(* IEC 61131-3 sources: PortalRobot/Portal_robot/Device/application/FB (part 4) *)

(* ---- FB_MAGAZINE.st ---- *)
FUNCTION_BLOCK FB_MAGAZINE
VAR_INPUT
	xIoManual : BOOL; // Передача выходов оператору отменяет пошаговую операцию
	uiMagazineId : UINT; // Идентификатор экземпляра 1..2
	xPointsConfigured : BOOL; // Настроена база этого магазина с Safe Z и Change Z
	xMechanismReady : BOOL := TRUE;
	xInventoryChanged : BOOL; // Сменился рабочий банк или оператор изменил его содержимое
	xTestInitialize : BOOL;
	xTestEnabled : BOOL;
	stRobotStatus     : ST_ROBOT_STATUS; // Текущие статусы робота
	astMachineStatus  : ARRAY [1..3] OF ST_MACHINE_PUBLIC; // Статусы станков для определения оставшейся работы
	auiMachineType    : ARRAY [1..3] OF UINT; // Тип детали, закреплённый за каждым станком
	stMagazineCommand : ST_MAGAZINE_COMMAND; // Команда магазина от автоматической логики
	stHmiCommand      : ST_ROBOT_COMMAND; // Ручная команда магазина с HMI
	xManual           : BOOL; // Разрешение ручного управления
	xReset            : BOOL; // Сброс ошибок магазина
	xResetCancel      : BOOL; // Отмена согласованного сброса по Stop/Disable
	RobotResetRecovery : ST_ROBOT_RESET_RECOVERY; // Внутреннее подтверждение принятого Reset робота
	xGlobalError      : BOOL; // Глобальная ошибка ячейки
	xHmiEnable        : BOOL; // Импульс включения магазина с HMI
	xHmiDisable       : BOOL; // Импульс отключения магазина с HMI
	xHmiFillBlanks    : BOOL; // Заполнить все активные слоты матрицы заготовками
	xHmiClear         : BOOL; // Полностью очистить содержимое магазина
	xHmiCycleSlot     : BOOL; // Переключить содержимое выбранного слота
	xHmiApplySlot     : BOOL; // Явно записать состояние и тип выбранного слота
	xHmiApplyPitchX   : BOOL; // Применить новый общий шаг слотов по X
	xHmiApplyPitchY   : BOOL; // Применить новый общий шаг слотов по Y
	uiHmiEditSlot     : UINT; // Номер слота для ручного редактирования
	uiHmiEditDetailType : UINT; // 0=NONE, 1=BLANK, 2=DETAIL
	uiHmiEditProductType : UINT; // Тип изделия 1..3
	lrHmiEditPitchX   : LREAL;
	lrHmiEditPitchY   : LREAL;
	xRobotOwnsMagazine : BOOL; // Автомат удерживает этот магазин в текущем цикле
	xRobotCanWorkWithMagazine : BOOL; // Интерфейс и точки готовы для роботной операции, не для включения магазина
	xSharedGeometryEditAllowed : BOOL; // Оба магазина выключены; общий шаг можно менять
	uiRows            : UINT; // Число строк матрицы магазина
	uiColumns         : UINT; // Число столбцов матрицы магазина
	uiTypeCount       : UINT; // Количество настроенных типов заготовок, 1..3
	auiSlotType       : ARRAY [1..GVL_CELL_SETTINGS.NumberDetail] OF UINT; // Тип секции каждого слота
	FaultRequest  : ST_MAGAZINE_FAULT_REQUEST; // Единый контракт диагностической инъекции
END_VAR
VAR_OUTPUT
    xInventoryUpdated : BOOL; // Только записи содержимого этим FB в текущем скане
	Command : ST_ROBOT_COMMAND; // Текущая пошаговая команда роботу
	Status  : ST_MAGAZINE_STATUS; // Рабочие статусы магазина
	Diag    : ST_MAGAZINE_DIAG; // Состояние автомата магазина
	Error   : ST_MAGAZINE_ERRORS; // Активные и последние ошибки
	FaultStatus : ST_FAULT_INJECTION_STATUS; // Состояние инжектора для HMI
END_VAR
VAR_IN_OUT
	stInventory : ST_MAGAZINE_INVENTORY; // Единственная кассета текущего магазина
	lrPitchX : LREAL; // Общий фактический шаг слотов по X
	lrPitchY : LREAL; // Общий фактический шаг слотов по Y
END_VAR
VAR
    xInventorySummaryInitialized : BOOL;
    xInventorySummaryDirty : BOOL;
    iInventorySummarySlotCount : SINT;
    uiInventorySummaryTypeCount : UINT;
    iInventoryFirstBlank : SINT;
    iInventoryFirstFree : SINT;
	eGrantedOperation : E_MAGAZINE_OPERATION; // Доступная операция магазина
	eActualOperation  : E_MAGAZINE_OPERATION; // Выполняемая операция магазина

	rtExecute          : R_TRIG; // Фронт команды запуска
	rtEnable           : R_TRIG; // Фронт команды включения
	rtDisable          : R_TRIG; // Фронт команды отключения
	rtFillBlanks       : R_TRIG; // Фронт заполнения магазина заготовками
	rtClear            : R_TRIG; // Фронт очистки магазина
	rtCycleSlot        : R_TRIG; // Фронт изменения выбранного слота
	rtApplySlot        : R_TRIG; // Фронт явной записи выбранного слота
	rtApplyPitchX      : R_TRIG;
	rtApplyPitchY      : R_TRIG;
	rtReset            : R_TRIG; // Фронт команды сброса магазина

	xExecuteRequest    : BOOL; // Активный запрос выполнения операции
	xResetRequest      : BOOL; // Активный запрос сброса
	xStopRequest       : BOOL; // Активный запрос остановки
	xManualCommand     : BOOL; // Команда получена из ручного интерфейса
	xDisableRequest    : BOOL; // Сохранённый запрос отключения после текущей операции
	xRobotInMagazineContext : BOOL; // Робот находится в рабочей зоне магазина
	xFaultContextCaptured : BOOL; // Контекст робота зафиксирован при входе в ERROR
	xRobotInMagazineAtFault : BOOL; // Робот был в рабочей зоне этого магазина при ошибке
	xRobotStopRequired : BOOL; // Итоговая реакция ROBOT_STOP, сформированная магазином
	xRobotResetDependencyReady : BOOL; // Каскадная ошибка робота может быть сброшена тем же импульсом
	xRobotResetDependencyRequired : BOOL; // Только ошибка с участием робота зависит от его восстановления
	xRobotResetCoordinated : BOOL; // Магазин присоединился к одному явно запрошенному сбросу
	udiRobotResetAttempt : UDINT; // Ожидаемый номер принятой попытки FB_ROBOT
	xRobotResetAttemptReady : BOOL; // Первичная зависимость восстановлена в той же попытке

	iActiveSlotCount   : SINT; // Число активных слотов выбранной матрицы
	iInventoryIndex    : SINT; // Индекс изменения содержимого магазина
	iTakeSlot          : SINT; // Слот выбранной заготовки
	iPutSlot           : SINT; // Выбранный свободный слот
	iActiveSlot        : SINT; // Единственный слот текущего элементарного движения
	xInventoryCommitted: BOOL; // Все изменения слотов текущей операции подтверждены
	xTakeSlotCommitted  : BOOL; // Изъятие заготовки отражено в матрице после закрытия захвата
	xPutSlotCommitted   : BOOL; // Укладка груза отражена в матрице после открытия захвата
	xRobotCommandStarted : BOOL; // Текущий элементарный шаг действительно принят FB_ROBOT
	xOperationSequenceComplete : BOOL; // Все шаги операции подтверждены до изменения матрицы
	xTakeSlotValid     : BOOL; // Проверка диапазона до обращения к массиву слотов
	xPutSlotValid      : BOOL;
	xTakeSlotHasBlank  : BOOL;
	xPutSlotEmpty      : BOOL;
	xChangeTakeFirst   : BOOL; // CHANGE в одном слоте: сначала TAKE, затем PUT
	xPutProductTypeValid : BOOL;
	uiStep             : UINT; // Шаг последовательности робота
	uiIndex            : UINT; // Индекс слота для расчёта координат

	stActiveRobotCommand : ST_ROBOT_COMMAND; // Команда роботу текущего шага
	xFinishedCondition   : BOOL; // Текущее содержимое не позволяет продолжить цикл
	xFinishedLatched     : BOOL; // Завершение этой палеты не отменяется работой другого магазина
	xMachineHasRelevantPart : BOOL; // В доступном станке есть заготовка, обработка или готовая деталь
	xMachineHasDestination : BOOL; // Для оставшейся работы есть свободный слот соответствующего типа
	xAllSlotsDetails    : BOOL; // Все активные слоты заполнены готовыми деталями
	xNoBlankNoMachinePart : BOOL; // Нет заготовок и нет доступной работы в станках
	xNoBlankNoDestination : BOOL; // Нет заготовок и нет места для возврата груза
	uiMachineIndex      : UINT; // Индекс станка при расчёте завершения магазина
	uiMachineTypeIndex  : UINT; // Тип детали проверяемого станка
	uiPutProductType    : UINT; // Тип груза, защёлкнутый до физического PUT
	fbFaultInjector      : FB_MAGAZINE_FAULT_INJECTOR; // Безопасный сценарий ошибки до движения
	xFaultAllowed        : BOOL; // Владелец разрешает синтетическую проверку
	xStartupInitialized  : BOOL;
	udiProducedPartsTotal : UDINT; // Монотонный счётчик подтверждённых укладок готовых деталей
END_VAR
VAR CONSTANT
	ERR_WRONG_OPERATION : DWORD := DWORD#16#0000_0001; // Недопустимая операция магазина
	ERR_NO_BLANK        : DWORD := DWORD#16#0000_0002; // В магазине нет заготовки
	ERR_NO_FREE_SLOT    : DWORD := DWORD#16#0000_0004; // В магазине нет свободного слота
	ERR_INVALID_SLOT    : DWORD := DWORD#16#0000_0008; // Недопустимый номер слота
	ERR_SLOT_CONTENT    : DWORD := DWORD#16#0000_0010; // Содержимое слота не соответствует операции
	ERR_ROBOT           : DWORD := DWORD#16#0000_0020; // Ошибка робота при операции магазина
	ERR_GLOBAL_STOP     : DWORD := DWORD#16#0000_0040; // Остановка по глобальной ошибке
	ERR_GEOMETRY        : DWORD := DWORD#16#0000_0080; // Ошибка параметров матрицы магазина
	MASK_EQUIPMENT_ERROR : DWORD := ERR_WRONG_OPERATION OR ERR_NO_BLANK
		OR ERR_NO_FREE_SLOT OR ERR_INVALID_SLOT OR ERR_SLOT_CONTENT OR ERR_GEOMETRY;
	WRN_RESET_EXECUTE_ACTIVE : UINT := 1; // Операция магазина ещё активна
	WRN_RESET_GLOBAL_ERROR   : UINT := 2; // Глобальная ошибка ещё активна
	WRN_RESET_ROBOT_ERROR    : UINT := 3; // Ошибка робота ещё активна
	WRN_ENABLE_GLOBAL_ERROR  : UINT := 4; // Включение запрещено глобальной ошибкой
	WRN_ENABLE_CONTENT       : UINT := 5; // Архив: содержимое больше не блокирует включение
	WRN_DISABLE_PENDING      : UINT := 6; // Отключение магазина уже запрошено
	WRN_FILL_ENABLED         : UINT := 7; // Заполнение запрещено для включённого магазина
	WRN_FILL_GEOMETRY        : UINT := 8; // Активная матрица магазина задана неверно
	WRN_CLEAR_ENABLED        : UINT := 9; // Очистка запрещена для включённого магазина
	WRN_SIM_ERROR_NOT_ALLOWED: UINT := 10; // Тестовая ошибка запрещена текущим состоянием
	WRN_EDIT_REJECTED : UINT := 14; // Редактирование включённого/занятого магазина запрещено
	WRN_GEOMETRY_EDIT_REJECTED : UINT := 16; // PLC отклонил изменение общего шага X/Y
	WRN_ENABLE_GEOMETRY      : UINT := 15; // Геометрия магазина не позволяет включение
	WRN_ENABLE_OWN_ERROR     : UINT := 17; // Включение запрещено собственной ошибкой магазина
	WRN_ENABLE_POINTS        : UINT := 18; // Не настроена база этого магазина или её Z-смещения
END_VAR

// --- BEGIN IMPLEMENTATION ---

xInventoryUpdated := FALSE;

// Инвентарь загружает владелец банков RunTwoPallet; здесь сбрасывается только автомат.
IF NOT xStartupInitialized THEN
	xFinishedLatched := FALSE;
	xFaultContextCaptured := FALSE;
	xRobotInMagazineAtFault := FALSE;
	xRobotStopRequired := FALSE;
	xStartupInitialized := TRUE;
END_IF;

IF xTestInitialize THEN
	xFinishedLatched := FALSE;
	IF xTestEnabled AND xPointsConfigured THEN
		Diag.eState := E_MAGAZINE_STATE.IDLE;
	ELSE
		Diag.eState := E_MAGAZINE_STATE.DISABLED;
	END_IF;
	Error.dwErrorActive := DWORD#0;
	Error.dwAlarmActive := DWORD#0;
	eGrantedOperation := E_MAGAZINE_OPERATION.NONE;
	eActualOperation := E_MAGAZINE_OPERATION.NONE;
	xExecuteRequest := FALSE;
	xResetRequest := FALSE;
	xStopRequest := FALSE;
	xManualCommand := FALSE;
	xDisableRequest := FALSE;
	iTakeSlot := SINT#0;
	iPutSlot := SINT#0;
	xChangeTakeFirst := FALSE;
	iActiveSlot := SINT#0;
	xInventoryCommitted := FALSE;
	xTakeSlotCommitted := FALSE;
	xPutSlotCommitted := FALSE;
	xRobotCommandStarted := FALSE;
	xOperationSequenceComplete := FALSE;
	xFaultContextCaptured := FALSE;
	xRobotInMagazineAtFault := FALSE;
	xRobotStopRequired := FALSE;
	uiStep := UINT#0;
	stActiveRobotCommand.xExecute := FALSE;
	stActiveRobotCommand.xStop := FALSE;
	stActiveRobotCommand.xReset := FALSE;
	stActiveRobotCommand.eAction := E_ROBOT_ACTION.NONE;
	stActiveRobotCommand.eSetPoint := E_POINT_NAME.NONE;
	stActiveRobotCommand.iActiveSlot := SINT#0;
	stActiveRobotCommand.uiMagazineId := uiMagazineId;
END_IF;

IF xInventoryChanged THEN
	xFinishedLatched := FALSE;
END_IF;

rtFillBlanks(CLK := xHmiFillBlanks);
rtClear(CLK := xHmiClear);
rtCycleSlot(CLK := xHmiCycleSlot);
rtApplySlot(CLK := xHmiApplySlot);
rtApplyPitchX(CLK := xHmiApplyPitchX);
rtApplyPitchY(CLK := xHmiApplyPitchY);

IF (uiRows > UINT#0)
AND (uiColumns > UINT#0)
AND ((uiRows * uiColumns) <= SINT_TO_UINT(GVL_CELL_SETTINGS.MagazineSlots)) THEN
	iActiveSlotCount := UINT_TO_SINT(uiRows * uiColumns);
ELSE
	iActiveSlotCount := SINT#0;
END_IF;

// Ручная роботная команда принадлежит только выбранному магазину.
xManualCommand := xManual
	AND (
		(stHmiCommand.eSetPoint = E_POINT_NAME.MAGAZINE_TAKE_DETAIL)
		OR (stHmiCommand.eSetPoint = E_POINT_NAME.MAGAZINE_PUT_DETAIL)
		OR (stHmiCommand.eSetPoint = E_POINT_NAME.MAGAZINE_CHANGE_DETAIL)
		OR (stHmiCommand.eSetPoint = E_POINT_NAME.MAGAZINE_RETURN_BLANK)
	)
	AND ((stHmiCommand.uiMagazineId = uiMagazineId)
		OR ((stHmiCommand.uiMagazineId = UINT#0) AND (uiMagazineId = UINT#1)));

IF xManual THEN
	IF xManualCommand THEN
		xExecuteRequest := stHmiCommand.xExecute;
		xStopRequest := stHmiCommand.xStop;
	ELSE
		xExecuteRequest := FALSE;
		xStopRequest := FALSE;
	END_IF;
ELSE
	xExecuteRequest := stMagazineCommand.xExecute;
	xStopRequest := stMagazineCommand.xStop;
END_IF;

// Контекст запрещает редактирование и завершает отложенное отключение только
// после фактического выхода робота из конкретного магазина.
xRobotInMagazineContext := (stRobotStatus.uiMagazineContext = uiMagazineId)
	OR ((stRobotStatus.uiMagazineContext = UINT#0)
		AND (xRobotOwnsMagazine OR xManualCommand)
		AND ((stRobotStatus.eCurrentPoint = E_POINT_NAME.MAGAZINE_IN_SLOT)
			OR (stRobotStatus.eCurrentPoint = E_POINT_NAME.MAGAZINE_CHANGE)));
xRobotInMagazineContext := xRobotInMagazineContext
	OR ((xRobotOwnsMagazine OR xManualCommand)
		AND (Diag.eState = E_MAGAZINE_STATE.ROBOT_COMMAND)
		AND (stActiveRobotCommand.eAction = E_ROBOT_ACTION.MOVE_TO_POINT)
		AND ((stActiveRobotCommand.eSetPoint = E_POINT_NAME.MAGAZINE_IN_SLOT)
			OR (stActiveRobotCommand.eSetPoint = E_POINT_NAME.MAGAZINE_CHANGE)));

// Единственную кассету можно менять только у технологически выключенного
// магазина, когда робот не находится внутри и не владеет текущей операцией.
Status.xEditAllowed := ((Diag.eState = E_MAGAZINE_STATE.DISABLED)
		OR (Diag.eState = E_MAGAZINE_STATE.ERROR))
	AND NOT xRobotOwnsMagazine
	AND NOT xRobotInMagazineContext
	AND NOT xGlobalError;
Status.xPitchEditAllowed := Status.xEditAllowed AND xSharedGeometryEditAllowed;

// Шаг матрицы общий для двух магазинов, поэтому менять его разрешено только
// когда оба магазина выключены. Смещения Z принадлежат базовым точкам магазина.
IF rtApplyPitchX.Q
AND Status.xEditAllowed
AND xSharedGeometryEditAllowed
AND (lrHmiEditPitchX >= LREAL#1.0)
AND (lrHmiEditPitchX <= LREAL#5000.0) THEN
	lrPitchX := lrHmiEditPitchX;
END_IF;
IF rtApplyPitchY.Q
AND Status.xEditAllowed
AND xSharedGeometryEditAllowed
AND (lrHmiEditPitchY >= LREAL#1.0)
AND (lrHmiEditPitchY <= LREAL#5000.0) THEN
	lrPitchY := lrHmiEditPitchY;
END_IF;
IF rtClear.Q AND Status.xEditAllowed THEN
	xFinishedLatched := FALSE;
	FOR iInventoryIndex := 1 TO GVL_CELL_SETTINGS.MagazineSlots DO
		xInventoryUpdated := TRUE;
		xInventorySummaryDirty := TRUE;
		stInventory.aSlots[iInventoryIndex].xInPosition := FALSE;
		stInventory.aSlots[iInventoryIndex].eDetailType := E_DETAIL_TYPE.NONE;
		stInventory.aSlots[iInventoryIndex].uiProductType := UINT#0;
	END_FOR;
ELSIF rtFillBlanks.Q
AND (iActiveSlotCount > SINT#0)
AND Status.xEditAllowed THEN
	xFinishedLatched := FALSE;
	FOR iInventoryIndex := 1 TO GVL_CELL_SETTINGS.MagazineSlots DO
		xInventoryUpdated := TRUE;
		xInventorySummaryDirty := TRUE;
		stInventory.aSlots[iInventoryIndex].xInPosition := iInventoryIndex <= iActiveSlotCount;
		IF iInventoryIndex <= iActiveSlotCount THEN
			stInventory.aSlots[iInventoryIndex].eDetailType := E_DETAIL_TYPE.BLANK;
			stInventory.aSlots[iInventoryIndex].uiProductType := auiSlotType[iInventoryIndex];
		ELSE
			stInventory.aSlots[iInventoryIndex].eDetailType := E_DETAIL_TYPE.NONE;
			stInventory.aSlots[iInventoryIndex].uiProductType := UINT#0;
		END_IF;
	END_FOR;
ELSIF rtApplySlot.Q
AND Status.xEditAllowed
AND (uiHmiEditSlot >= UINT#1)
AND (uiHmiEditSlot <= SINT_TO_UINT(iActiveSlotCount))
AND (uiHmiEditDetailType <= UINT#2)
AND ((uiHmiEditDetailType = UINT#0)
	OR ((uiHmiEditProductType >= UINT#1) AND (uiHmiEditProductType <= uiTypeCount))) THEN
	xFinishedLatched := FALSE;
	iInventoryIndex := UINT_TO_SINT(uiHmiEditSlot);
	CASE uiHmiEditDetailType OF
		UINT#0:
			xInventoryUpdated := TRUE;
			xInventorySummaryDirty := TRUE;
			stInventory.aSlots[iInventoryIndex].xInPosition := FALSE;
			stInventory.aSlots[iInventoryIndex].eDetailType := E_DETAIL_TYPE.NONE;
			stInventory.aSlots[iInventoryIndex].uiProductType := UINT#0;
		UINT#1:
			xInventoryUpdated := TRUE;
			xInventorySummaryDirty := TRUE;
			stInventory.aSlots[iInventoryIndex].xInPosition := TRUE;
			stInventory.aSlots[iInventoryIndex].eDetailType := E_DETAIL_TYPE.BLANK;
			stInventory.aSlots[iInventoryIndex].uiProductType := uiHmiEditProductType;
		UINT#2:
			xInventoryUpdated := TRUE;
			xInventorySummaryDirty := TRUE;
			stInventory.aSlots[iInventoryIndex].xInPosition := TRUE;
			stInventory.aSlots[iInventoryIndex].eDetailType := E_DETAIL_TYPE.DETAIL;
			stInventory.aSlots[iInventoryIndex].uiProductType := uiHmiEditProductType;
	END_CASE;
ELSIF rtCycleSlot.Q
AND Status.xEditAllowed
AND (uiHmiEditSlot >= UINT#1)
AND (uiHmiEditSlot <= SINT_TO_UINT(iActiveSlotCount)) THEN
	xFinishedLatched := FALSE;
	iInventoryIndex := UINT_TO_SINT(uiHmiEditSlot);
	IF NOT stInventory.aSlots[iInventoryIndex].xInPosition
	OR (stInventory.aSlots[iInventoryIndex].eDetailType = E_DETAIL_TYPE.NONE) THEN
		xInventoryUpdated := TRUE;
		xInventorySummaryDirty := TRUE;
		stInventory.aSlots[iInventoryIndex].xInPosition := TRUE;
		stInventory.aSlots[iInventoryIndex].eDetailType := E_DETAIL_TYPE.BLANK;
		stInventory.aSlots[iInventoryIndex].uiProductType := auiSlotType[iInventoryIndex];
	ELSE
		xInventoryUpdated := TRUE;
		xInventorySummaryDirty := TRUE;
		stInventory.aSlots[iInventoryIndex].xInPosition := FALSE;
		stInventory.aSlots[iInventoryIndex].eDetailType := E_DETAIL_TYPE.NONE;
		stInventory.aSlots[iInventoryIndex].uiProductType := UINT#0;
	END_IF;
END_IF;

// При смене банка проверка завершения использует его текущую карту типов,
// а не свободные слоты прежней палеты с прошлого скана.
IF NOT xInventorySummaryInitialized OR xInventoryChanged OR xTestInitialize
OR (iInventorySummarySlotCount <> iActiveSlotCount)
OR (uiInventorySummaryTypeCount <> uiTypeCount) THEN
    xInventorySummaryDirty := TRUE;
END_IF;
IF xInventorySummaryDirty THEN
    UpdateTypeStatus(stMagazineInventory := stInventory);
END_IF;
Status.iCurrentBlank := iInventoryFirstBlank;
Status.iCurrentFreeSlot := iInventoryFirstFree;

Status.xOutBlank := Status.iCurrentBlank = SINT#0;
Status.xOutFreeSlot := Status.iCurrentFreeSlot = SINT#0;
Status.xCanTake := NOT Status.xOutBlank;
Status.xCanPut := NOT Status.xOutFreeSlot;
Status.xCanChange := Status.xCanTake; // Изъятие заготовки само освобождает место
Status.xCanEnable := FALSE;

// Для PUT/возврата заготовки нужен пустой слот. Готовую деталь можно обменять
// на заготовку в одном занятом слоте, если первый захват свободен и открыт.
IF stRobotStatus.xBlankAvailable OR stRobotStatus.xDetailAvailable THEN
	Status.xCanEnable := Status.xCanPut;
ELSIF NOT stRobotStatus.xBlankAvailable AND NOT stRobotStatus.xDetailAvailable THEN
	Status.xCanEnable := Status.xCanTake;
END_IF;

IF stRobotStatus.xDetailAvailable AND NOT stRobotStatus.xBlankAvailable
AND stRobotStatus.xGripper1Open AND Status.xCanChange THEN
	Status.xCanEnable := TRUE;
END_IF;

// Отсутствие заготовок не завершает магазин, пока из станков ещё можно вернуть
// готовую деталь в свободный слот соответствующего типа.
xMachineHasRelevantPart := FALSE;
xMachineHasDestination := FALSE;
FOR uiMachineIndex := UINT#1 TO UINT#3 DO
	IF astMachineStatus[uiMachineIndex].xEnabled
	AND NOT astMachineStatus[uiMachineIndex].xError
	AND (astMachineStatus[uiMachineIndex].xProcessing
		OR ((astMachineStatus[uiMachineIndex].ePartState = E_PART_STATE.LOADED)
			AND ((astMachineStatus[uiMachineIndex].ePartType = E_PART_TYPE.PART)
				OR (astMachineStatus[uiMachineIndex].ePartType = E_PART_TYPE.DETAIL)))) THEN
		xMachineHasRelevantPart := TRUE;
		uiMachineTypeIndex := auiMachineType[uiMachineIndex];
		IF (uiMachineTypeIndex >= UINT#1)
		AND (uiMachineTypeIndex <= UINT#3)
		AND (Status.stTypeStatus.aiFreeSlot[uiMachineTypeIndex] > SINT#0) THEN
			xMachineHasDestination := TRUE;
		END_IF;
	END_IF;
END_FOR;

IF NOT stRobotStatus.xBlankAvailable
AND NOT stRobotStatus.xDetailAvailable
AND xMachineHasDestination THEN
	Status.xCanEnable := TRUE;
END_IF;

Status.xEnableCheckRobotReady := xRobotCanWorkWithMagazine AND xMechanismReady;
Status.xEnableCheckRobotReleased := NOT xRobotInMagazineContext;
Status.xEnableCheckNoError := NOT xGlobalError
	AND (Diag.eState <> E_MAGAZINE_STATE.ERROR)
	AND (Error.dwErrorActive = DWORD#0);
Status.xEnableCheckContent := Status.xCanEnable;
Status.xEnableCheckGeometry := (iActiveSlotCount > SINT#0)
	AND (lrPitchX >= LREAL#1.0)
	AND (lrPitchX <= LREAL#5000.0)
	AND (lrPitchY >= LREAL#1.0)
	AND (lrPitchY <= LREAL#5000.0);
// Включение требует собственную базовую точку магазина. Готовность интерфейса,
// положение робота и содержимое палеты проверяются при роботной операции.
Status.xEnableSequenceAllowed := (Diag.eState = E_MAGAZINE_STATE.DISABLED)
	AND Status.xEnableCheckNoError
	AND Status.xEnableCheckGeometry
	AND xPointsConfigured;

// Finished остаётся прежним по смыслу, но теперь оценивает единственную кассету.
xAllSlotsDetails := iActiveSlotCount > SINT#0;
IF xAllSlotsDetails THEN
	FOR uiIndex := UINT#1 TO SINT_TO_UINT(iActiveSlotCount) DO
		IF NOT stInventory.aSlots[UINT_TO_SINT(uiIndex)].xInPosition
		OR (stInventory.aSlots[UINT_TO_SINT(uiIndex)].eDetailType <> E_DETAIL_TYPE.DETAIL) THEN
			xAllSlotsDetails := FALSE;
		END_IF;
	END_FOR;
END_IF;
xNoBlankNoMachinePart := Status.xOutBlank AND NOT xMachineHasRelevantPart;
xNoBlankNoDestination := Status.xOutBlank AND NOT xMachineHasDestination;
xFinishedCondition :=
	(NOT stRobotStatus.xBlankAvailable AND NOT stRobotStatus.xDetailAvailable)
	AND (xAllSlotsDetails OR xNoBlankNoMachinePart OR xNoBlankNoDestination);

eGrantedOperation := E_MAGAZINE_OPERATION.NONE;
IF stRobotStatus.xBlankAvailable
AND stRobotStatus.xDetailAvailable
AND Status.xCanPut THEN
	// Сначала освобождается захват готовой детали; заготовка остаётся у робота.
	eGrantedOperation := E_MAGAZINE_OPERATION.PUT;
ELSIF NOT Status.xOutBlank
AND NOT stRobotStatus.xBlankAvailable
AND NOT stRobotStatus.xDetailAvailable THEN
	eGrantedOperation := E_MAGAZINE_OPERATION.TAKE;
ELSIF NOT Status.xOutBlank
AND stRobotStatus.xGripper1Open
AND NOT stRobotStatus.xBlankAvailable
AND stRobotStatus.xDetailAvailable THEN
	eGrantedOperation := E_MAGAZINE_OPERATION.CHANGE;
ELSIF NOT Status.xOutFreeSlot
AND stRobotStatus.xDetailAvailable THEN
	eGrantedOperation := E_MAGAZINE_OPERATION.PUT;
END_IF;

xResetRequest := xReset;
rtReset(CLK := xResetRequest);

// RunMagazine предшествует RunRobot. В скане нажатия ожидаем следующий номер;
// на следующем скане уже требуется подтверждённая, всё ещё активная попытка.
IF xRobotResetCoordinated
AND (NOT RobotResetRecovery.xActive
	OR (RobotResetRecovery.udiAttempt <> udiRobotResetAttempt)
	OR xGlobalError OR xIoManual OR xStopRequest OR xExecuteRequest OR xResetCancel) THEN
	xRobotResetCoordinated := FALSE;
	IF (Diag.eState = E_MAGAZINE_STATE.ERROR) AND stRobotStatus.xError THEN
		Diag.stWarning.uiCode := WRN_RESET_ROBOT_ERROR;
		Diag.stWarning.udiSequence := Diag.stWarning.udiSequence + UDINT#1;
		IF Diag.stWarning.udiSequence = UDINT#0 THEN Diag.stWarning.udiSequence := UDINT#1; END_IF;
	END_IF;
END_IF;
xRobotResetAttemptReady := xRobotResetCoordinated
	AND RobotResetRecovery.xActive
	AND (RobotResetRecovery.udiAttempt = udiRobotResetAttempt)
	AND RobotResetRecovery.xDependenciesReady;

xRobotResetDependencyRequired := ((Error.dwErrorActive AND ERR_ROBOT) <> DWORD#0)
	OR xRobotInMagazineAtFault;
xRobotResetDependencyReady := NOT xRobotResetDependencyRequired
	OR NOT stRobotStatus.xError
	OR stRobotStatus.xResetAllowed
	OR xRobotResetAttemptReady;

IF rtReset.Q
AND (Diag.eState = E_MAGAZINE_STATE.ERROR) THEN
	IF xExecuteRequest THEN
		Diag.stWarning.uiCode := WRN_RESET_EXECUTE_ACTIVE;
	ELSIF xGlobalError THEN
		Diag.stWarning.uiCode := WRN_RESET_GLOBAL_ERROR;
	ELSIF stRobotStatus.xError
	AND NOT stRobotStatus.xResetAllowed THEN
		Diag.stWarning.uiCode := WRN_RESET_ROBOT_ERROR;
	ELSE
		Diag.stWarning.uiCode := UINT#0;
	END_IF;

	IF Diag.stWarning.uiCode <> UINT#0 THEN
		Diag.stWarning.udiSequence := Diag.stWarning.udiSequence + UDINT#1;
		IF Diag.stWarning.udiSequence = UDINT#0 THEN
			Diag.stWarning.udiSequence := UDINT#1;
		END_IF;
	END_IF;
END_IF;

rtEnable(CLK := xHmiEnable OR (NOT xManual AND stMagazineCommand.xEnable));
rtDisable(CLK := xHmiDisable OR (NOT xManual AND stMagazineCommand.xDisable));

IF rtEnable.Q
AND (Diag.eState = E_MAGAZINE_STATE.DISABLED)
AND NOT Status.xEnableSequenceAllowed THEN
	IF NOT xPointsConfigured THEN
		Diag.stWarning.uiCode := WRN_ENABLE_POINTS;
	ELSIF xGlobalError THEN
		Diag.stWarning.uiCode := WRN_ENABLE_GLOBAL_ERROR;
	ELSIF NOT Status.xEnableCheckGeometry THEN
		Diag.stWarning.uiCode := WRN_ENABLE_GEOMETRY;
	ELSE
		Diag.stWarning.uiCode := WRN_ENABLE_OWN_ERROR;
	END_IF;
	Diag.stWarning.udiSequence := Diag.stWarning.udiSequence + UDINT#1;
	IF Diag.stWarning.udiSequence = UDINT#0 THEN
		Diag.stWarning.udiSequence := UDINT#1;
	END_IF;
ELSIF rtDisable.Q
AND xHmiDisable
AND xDisableRequest THEN
	Diag.stWarning.uiCode := WRN_DISABLE_PENDING;
	Diag.stWarning.udiSequence := Diag.stWarning.udiSequence + UDINT#1;
	IF Diag.stWarning.udiSequence = UDINT#0 THEN
		Diag.stWarning.udiSequence := UDINT#1;
	END_IF;
ELSIF rtFillBlanks.Q
AND (iActiveSlotCount = 0) THEN
	Diag.stWarning.uiCode := WRN_FILL_GEOMETRY;
	Diag.stWarning.udiSequence := Diag.stWarning.udiSequence + UDINT#1;
	IF Diag.stWarning.udiSequence = UDINT#0 THEN
		Diag.stWarning.udiSequence := UDINT#1;
	END_IF;
ELSIF rtFillBlanks.Q
AND NOT Status.xEditAllowed THEN
	Diag.stWarning.uiCode := WRN_FILL_ENABLED;
	Diag.stWarning.udiSequence := Diag.stWarning.udiSequence + UDINT#1;
	IF Diag.stWarning.udiSequence = UDINT#0 THEN
		Diag.stWarning.udiSequence := UDINT#1;
	END_IF;
ELSIF rtClear.Q
AND NOT Status.xEditAllowed THEN
	Diag.stWarning.uiCode := WRN_CLEAR_ENABLED;
	Diag.stWarning.udiSequence := Diag.stWarning.udiSequence + UDINT#1;
	IF Diag.stWarning.udiSequence = UDINT#0 THEN
		Diag.stWarning.udiSequence := UDINT#1;
	END_IF;
ELSIF (rtApplyPitchX.Q
	AND (NOT Status.xEditAllowed
		OR NOT xSharedGeometryEditAllowed
		OR (lrHmiEditPitchX < LREAL#1.0)
		OR (lrHmiEditPitchX > LREAL#5000.0)))
OR (rtApplyPitchY.Q
	AND (NOT Status.xEditAllowed
		OR NOT xSharedGeometryEditAllowed
		OR (lrHmiEditPitchY < LREAL#1.0)
		OR (lrHmiEditPitchY > LREAL#5000.0))) THEN
	Diag.stWarning.uiCode := WRN_GEOMETRY_EDIT_REJECTED;
	Diag.stWarning.udiSequence := Diag.stWarning.udiSequence + UDINT#1;
	IF Diag.stWarning.udiSequence = UDINT#0 THEN
		Diag.stWarning.udiSequence := UDINT#1;
	END_IF;
ELSIF rtApplySlot.Q
AND ((uiHmiEditSlot < UINT#1)
	OR (uiHmiEditSlot > SINT_TO_UINT(iActiveSlotCount))
	OR (uiHmiEditDetailType > UINT#2)
	OR ((uiHmiEditDetailType <> UINT#0)
		AND ((uiHmiEditProductType < UINT#1) OR (uiHmiEditProductType > uiTypeCount)))
	OR NOT Status.xEditAllowed) THEN
	Diag.stWarning.uiCode := WRN_EDIT_REJECTED;
	Diag.stWarning.udiSequence := Diag.stWarning.udiSequence + UDINT#1;
	IF Diag.stWarning.udiSequence = UDINT#0 THEN
		Diag.stWarning.udiSequence := UDINT#1;
	END_IF;
ELSIF rtCycleSlot.Q
AND ((uiHmiEditSlot < UINT#1)
	OR (uiHmiEditSlot > SINT_TO_UINT(iActiveSlotCount))
	OR NOT Status.xEditAllowed) THEN
	Diag.stWarning.uiCode := WRN_EDIT_REJECTED;
	Diag.stWarning.udiSequence := Diag.stWarning.udiSequence + UDINT#1;
	IF Diag.stWarning.udiSequence = UDINT#0 THEN
		Diag.stWarning.udiSequence := UDINT#1;
	END_IF;
END_IF;

IF rtDisable.Q THEN
	xDisableRequest := TRUE;
END_IF;

rtExecute(CLK := xExecuteRequest);

// Синтетический сценарий входит только в проверочный шаг CHOOSE и не выдаёт
// команду движения роботу до формирования выбранной штатной ошибки.
xFaultAllowed := ((Diag.eState = E_MAGAZINE_STATE.DISABLED)
	OR (Diag.eState = E_MAGAZINE_STATE.IDLE))
	AND NOT xExecuteRequest
	AND NOT xGlobalError
	AND NOT stRobotStatus.xBusy
	AND NOT stRobotStatus.xError
	AND (Error.dwErrorActive = DWORD#0);

fbFaultInjector(
	Request := FaultRequest,
	xOwnerAllowed := xFaultAllowed,
	xComplete := Diag.eState = E_MAGAZINE_STATE.ERROR
);
FaultStatus := fbFaultInjector.Status;

IF fbFaultInjector.Status.xRejected THEN
	Diag.stWarning.uiCode := WRN_SIM_ERROR_NOT_ALLOWED;
	Diag.stWarning.udiSequence := Diag.stWarning.udiSequence + UDINT#1;
	IF Diag.stWarning.udiSequence = UDINT#0 THEN
		Diag.stWarning.udiSequence := UDINT#1;
	END_IF;
END_IF;

// Значения команды роботу по умолчанию.
Command.xExecute := FALSE;
Command.xStop := FALSE;
Command.xReset := xResetRequest;
Command.eAction := E_ROBOT_ACTION.NONE;
Command.eSetPoint := E_POINT_NAME.NONE;
Command.iActiveSlot := 0;
Command.uiMagazineId := UINT#0;

// Ошибка робота в рабочей зоне принадлежит одновременно роботу и магазину.
IF xRobotInMagazineContext
AND stRobotStatus.xError
AND NOT xRobotResetAttemptReady
AND (Diag.eState <> E_MAGAZINE_STATE.ERROR) THEN
	Error.dwErrorActive := Error.dwErrorActive OR ERR_ROBOT;
	Diag.eState := E_MAGAZINE_STATE.ERROR;
END_IF;

IF xGlobalError
AND (Diag.eState <> E_MAGAZINE_STATE.DISABLED)
AND (Diag.eState <> E_MAGAZINE_STATE.IDLE)
AND (Diag.eState <> E_MAGAZINE_STATE.ERROR) THEN
	Error.dwErrorActive := Error.dwErrorActive OR ERR_GLOBAL_STOP;
	Diag.eState := E_MAGAZINE_STATE.ERROR;
END_IF;

// Сохраняем уже подтверждённые изменения слотов и первичную аварию,
// но не оставляем команду, которая продолжится после возврата I/O программе.
IF xIoManual THEN
	xExecuteRequest := FALSE;
	xStopRequest := FALSE;
	xDisableRequest := FALSE;
	xRobotCommandStarted := FALSE;
	xOperationSequenceComplete := FALSE;
	eActualOperation := E_MAGAZINE_OPERATION.NONE;
	stActiveRobotCommand.xExecute := FALSE;
	IF Diag.eState <> E_MAGAZINE_STATE.ERROR THEN
		Diag.eState := E_MAGAZINE_STATE.DISABLED;
	END_IF;
END_IF;

CASE Diag.eState OF
	E_MAGAZINE_STATE.DISABLED:
		xDisableRequest := FALSE;
		IF fbFaultInjector.Status.xBusy THEN
			iTakeSlot := 1;
			iPutSlot := 1;
			IF fbFaultInjector.xWrongOperation THEN
				eActualOperation := E_MAGAZINE_OPERATION.NONE;
			ELSIF fbFaultInjector.xNoFreeSlot THEN
				eActualOperation := E_MAGAZINE_OPERATION.PUT;
			ELSE
				eActualOperation := E_MAGAZINE_OPERATION.TAKE;
			END_IF;
			Diag.eState := E_MAGAZINE_STATE.CHOOSE;
		ELSIF rtEnable.Q AND NOT xIoManual
		AND Status.xEnableSequenceAllowed THEN
			Diag.eState := E_MAGAZINE_STATE.IDLE;
		END_IF;

	E_MAGAZINE_STATE.IDLE:
		uiStep := 0;
		eActualOperation := E_MAGAZINE_OPERATION.NONE;
		xInventoryCommitted := FALSE;
		xTakeSlotCommitted := FALSE;
		xPutSlotCommitted := FALSE;
		xOperationSequenceComplete := FALSE;

		IF fbFaultInjector.Status.xBusy THEN
			iTakeSlot := 1;
			iPutSlot := 1;
			IF fbFaultInjector.xWrongOperation THEN
				eActualOperation := E_MAGAZINE_OPERATION.NONE;
			ELSIF fbFaultInjector.xNoFreeSlot THEN
				eActualOperation := E_MAGAZINE_OPERATION.PUT;
			ELSE
				eActualOperation := E_MAGAZINE_OPERATION.TAKE;
			END_IF;
			Diag.eState := E_MAGAZINE_STATE.CHOOSE;
		ELSIF xFinishedLatched OR xFinishedCondition THEN
			Diag.eState := E_MAGAZINE_STATE.DISABLED;
		// Активный автоматический цикл сначала должен передать владение второму
		// магазину. До этого сохраняем xEnabled + xDisablePending, иначе менеджер
		// остаётся владельцем уже выключенного магазина и не может продолжить груз.
		ELSIF xDisableRequest
		AND NOT xRobotInMagazineContext THEN
			Diag.eState := E_MAGAZINE_STATE.DISABLED;
		ELSIF xGlobalError THEN
			Error.dwErrorActive := Error.dwErrorActive OR ERR_GLOBAL_STOP;
			Diag.eState := E_MAGAZINE_STATE.ERROR;
		// Автоматический владелец держит xExecute до завершения операции. Если
		// команда пришла раньше включения магазина, фронт был бы поглощён в
		// DISABLED; в IDLE принимаем также активный уровень запроса.
		ELSIF (rtExecute.Q OR xExecuteRequest) AND xMechanismReady THEN
			IF xManualCommand THEN
				CASE stHmiCommand.eSetPoint OF
					E_POINT_NAME.MAGAZINE_TAKE_DETAIL:
						eActualOperation := E_MAGAZINE_OPERATION.TAKE;
						iTakeSlot := stHmiCommand.iActiveSlot;
					E_POINT_NAME.MAGAZINE_PUT_DETAIL:
						eActualOperation := E_MAGAZINE_OPERATION.PUT;
						iPutSlot := stHmiCommand.iActiveSlot;
					E_POINT_NAME.MAGAZINE_CHANGE_DETAIL:
						// CHANGE требует двух слотов и запускается через ST_MAGAZINE_COMMAND.
						eActualOperation := E_MAGAZINE_OPERATION.NONE;
					E_POINT_NAME.MAGAZINE_RETURN_BLANK:
						eActualOperation := E_MAGAZINE_OPERATION.RETURN_BLANK;
						iPutSlot := stHmiCommand.iActiveSlot;
				ELSE
						eActualOperation := E_MAGAZINE_OPERATION.NONE;
				END_CASE;
			ELSE
				eActualOperation := stMagazineCommand.eOperation;
				iTakeSlot := stMagazineCommand.iTakeSlot;
				iPutSlot := stMagazineCommand.iPutSlot;
			END_IF;

			Diag.eState := E_MAGAZINE_STATE.CHOOSE;
		END_IF;

	E_MAGAZINE_STATE.CHOOSE:
		xTakeSlotValid := (iTakeSlot >= 1) AND (iTakeSlot <= iActiveSlotCount);
		xPutSlotValid := (iPutSlot >= 1) AND (iPutSlot <= iActiveSlotCount);
		xChangeTakeFirst := (eActualOperation = E_MAGAZINE_OPERATION.CHANGE)
			AND (iTakeSlot = iPutSlot);
		xTakeSlotHasBlank := FALSE;
		xPutSlotEmpty := FALSE;

		IF xTakeSlotValid THEN
		xTakeSlotHasBlank := stInventory.aSlots[iTakeSlot].xInPosition
			AND (stInventory.aSlots[iTakeSlot].eDetailType = E_DETAIL_TYPE.BLANK)
			AND (stInventory.aSlots[iTakeSlot].uiProductType >= UINT#1)
			AND (stInventory.aSlots[iTakeSlot].uiProductType <= uiTypeCount);
		END_IF;

	IF xPutSlotValid THEN
		xPutSlotEmpty := NOT stInventory.aSlots[iPutSlot].xInPosition;
	END_IF;
	xPutProductTypeValid := TRUE;
	IF (eActualOperation = E_MAGAZINE_OPERATION.PUT)
	OR (eActualOperation = E_MAGAZINE_OPERATION.CHANGE) THEN
		xPutProductTypeValid := (stRobotStatus.uiDetailPayloadType >= UINT#1)
			AND (stRobotStatus.uiDetailPayloadType <= uiTypeCount);
	ELSIF eActualOperation = E_MAGAZINE_OPERATION.RETURN_BLANK THEN
		xPutProductTypeValid := (stRobotStatus.uiBlankPayloadType >= UINT#1)
			AND (stRobotStatus.uiBlankPayloadType <= uiTypeCount);
	END_IF;

		IF fbFaultInjector.xGeometry
		OR (iActiveSlotCount = 0) THEN
			Error.dwErrorActive := Error.dwErrorActive OR ERR_GEOMETRY;
			Diag.eState := E_MAGAZINE_STATE.ERROR;

		ELSIF fbFaultInjector.xWrongOperation
		OR (eActualOperation = E_MAGAZINE_OPERATION.NONE) THEN
			Error.dwErrorActive := Error.dwErrorActive OR ERR_WRONG_OPERATION;
			Diag.eState := E_MAGAZINE_STATE.ERROR;

		ELSIF fbFaultInjector.xNoBlank THEN
			Error.dwErrorActive := Error.dwErrorActive OR ERR_NO_BLANK;
			Diag.eState := E_MAGAZINE_STATE.ERROR;

		ELSIF fbFaultInjector.xNoFreeSlot THEN
			Error.dwErrorActive := Error.dwErrorActive OR ERR_NO_FREE_SLOT;
			Diag.eState := E_MAGAZINE_STATE.ERROR;

		ELSIF fbFaultInjector.xInvalidSlot THEN
			Error.dwErrorActive := Error.dwErrorActive OR ERR_INVALID_SLOT;
			Diag.eState := E_MAGAZINE_STATE.ERROR;

		ELSIF fbFaultInjector.xSlotContent THEN
			Error.dwErrorActive := Error.dwErrorActive OR ERR_SLOT_CONTENT;
			Diag.eState := E_MAGAZINE_STATE.ERROR;

		ELSIF ((eActualOperation = E_MAGAZINE_OPERATION.TAKE)
			OR (eActualOperation = E_MAGAZINE_OPERATION.CHANGE))
		AND NOT xTakeSlotValid THEN
			Error.dwErrorActive := Error.dwErrorActive OR ERR_NO_BLANK OR ERR_INVALID_SLOT;
			Diag.eState := E_MAGAZINE_STATE.ERROR;

		ELSIF ((eActualOperation = E_MAGAZINE_OPERATION.PUT)
			OR (eActualOperation = E_MAGAZINE_OPERATION.CHANGE)
			OR (eActualOperation = E_MAGAZINE_OPERATION.RETURN_BLANK))
		AND NOT xPutSlotValid THEN
			Error.dwErrorActive := Error.dwErrorActive OR ERR_NO_FREE_SLOT OR ERR_INVALID_SLOT;
			Diag.eState := E_MAGAZINE_STATE.ERROR;

		ELSIF ((eActualOperation = E_MAGAZINE_OPERATION.TAKE)
			OR (eActualOperation = E_MAGAZINE_OPERATION.CHANGE))
		AND NOT xTakeSlotHasBlank THEN
			Error.dwErrorActive := Error.dwErrorActive OR ERR_SLOT_CONTENT;
			Diag.eState := E_MAGAZINE_STATE.ERROR;

		ELSIF ((eActualOperation = E_MAGAZINE_OPERATION.PUT)
			OR (eActualOperation = E_MAGAZINE_OPERATION.CHANGE)
			OR (eActualOperation = E_MAGAZINE_OPERATION.RETURN_BLANK))
		AND NOT xPutSlotEmpty
		AND NOT (xChangeTakeFirst AND xTakeSlotHasBlank) THEN
			Error.dwErrorActive := Error.dwErrorActive OR ERR_SLOT_CONTENT;
			Diag.eState := E_MAGAZINE_STATE.ERROR;

		ELSIF ((eActualOperation = E_MAGAZINE_OPERATION.PUT)
			OR (eActualOperation = E_MAGAZINE_OPERATION.CHANGE)
			OR (eActualOperation = E_MAGAZINE_OPERATION.RETURN_BLANK))
		AND NOT xPutProductTypeValid THEN
			Error.dwErrorActive := Error.dwErrorActive OR ERR_SLOT_CONTENT;
			Diag.eState := E_MAGAZINE_STATE.ERROR;

		ELSIF (eActualOperation = E_MAGAZINE_OPERATION.TAKE)
		AND (stRobotStatus.xBlankAvailable OR stRobotStatus.xDetailAvailable) THEN
			Error.dwErrorActive := Error.dwErrorActive OR ERR_WRONG_OPERATION;
			Diag.eState := E_MAGAZINE_STATE.ERROR;

		ELSIF (eActualOperation = E_MAGAZINE_OPERATION.CHANGE)
		AND (NOT stRobotStatus.xGripper1Open
			OR stRobotStatus.xBlankAvailable) THEN
			Error.dwErrorActive := Error.dwErrorActive OR ERR_WRONG_OPERATION;
			Diag.eState := E_MAGAZINE_STATE.ERROR;

		ELSIF ((eActualOperation = E_MAGAZINE_OPERATION.PUT)
			OR (eActualOperation = E_MAGAZINE_OPERATION.CHANGE))
		AND NOT stRobotStatus.xDetailAvailable THEN
			Error.dwErrorActive := Error.dwErrorActive OR ERR_WRONG_OPERATION;
			Diag.eState := E_MAGAZINE_STATE.ERROR;

		ELSIF (eActualOperation = E_MAGAZINE_OPERATION.RETURN_BLANK)
		AND (NOT stRobotStatus.xBlankAvailable
			OR stRobotStatus.xDetailAvailable) THEN
			Error.dwErrorActive := Error.dwErrorActive OR ERR_WRONG_OPERATION;
			Diag.eState := E_MAGAZINE_STATE.ERROR;

		ELSE
			uiPutProductType := UINT#0;
			IF (eActualOperation = E_MAGAZINE_OPERATION.PUT)
			OR (eActualOperation = E_MAGAZINE_OPERATION.CHANGE) THEN
				uiPutProductType := stRobotStatus.uiDetailPayloadType;
			ELSIF eActualOperation = E_MAGAZINE_OPERATION.RETURN_BLANK THEN
				uiPutProductType := stRobotStatus.uiBlankPayloadType;
			END_IF;
			xInventoryCommitted := FALSE;
			xTakeSlotCommitted := FALSE;
			xPutSlotCommitted := FALSE;
			xOperationSequenceComplete := FALSE;
			uiStep := 0;
			Diag.eState := E_MAGAZINE_STATE.PREPARE_STEP;
		END_IF;

	E_MAGAZINE_STATE.PREPARE_STEP:
		xRobotCommandStarted := FALSE;
		stActiveRobotCommand.xExecute := FALSE;
		stActiveRobotCommand.xStop := FALSE;
		stActiveRobotCommand.xReset := xResetRequest;
		stActiveRobotCommand.eAction := E_ROBOT_ACTION.NONE;
		stActiveRobotCommand.eSetPoint := E_POINT_NAME.NONE;

		CASE eActualOperation OF
			E_MAGAZINE_OPERATION.TAKE:
				iActiveSlot := iTakeSlot;
			E_MAGAZINE_OPERATION.PUT,
			E_MAGAZINE_OPERATION.RETURN_BLANK:
				iActiveSlot := iPutSlot;
			E_MAGAZINE_OPERATION.CHANGE:
				IF uiStep <= UINT#5 THEN
					iActiveSlot := iPutSlot;
				ELSE
					iActiveSlot := iTakeSlot;
				END_IF;
		ELSE
			iActiveSlot := SINT#0;
		END_CASE;
		stActiveRobotCommand.iActiveSlot := iActiveSlot;
		stActiveRobotCommand.uiMagazineId := uiMagazineId;

		CASE eActualOperation OF
				E_MAGAZINE_OPERATION.TAKE:
					CASE uiStep OF
						0:
							IF stRobotStatus.xRotatedToDetail THEN
								Diag.eState := E_MAGAZINE_STATE.NEXT;
							ELSE
								stActiveRobotCommand.eAction := E_ROBOT_ACTION.ROTATE_TO_DETAIL;
							END_IF;
						1:
							stActiveRobotCommand.eAction := E_ROBOT_ACTION.MOVE_TO_POINT;
							stActiveRobotCommand.eSetPoint := E_POINT_NAME.MAGAZINE_SAFE;
						2:
							stActiveRobotCommand.eAction := E_ROBOT_ACTION.MOVE_TO_POINT;
							stActiveRobotCommand.eSetPoint := E_POINT_NAME.MAGAZINE_IN_SLOT;
						3: stActiveRobotCommand.eAction := E_ROBOT_ACTION.CLAMP_1;
						4:
							stActiveRobotCommand.eAction := E_ROBOT_ACTION.MOVE_TO_POINT;
							stActiveRobotCommand.eSetPoint := E_POINT_NAME.MAGAZINE_SAFE;
					ELSE
						xOperationSequenceComplete := TRUE;
						Diag.eState := E_MAGAZINE_STATE.DONE;
					END_CASE;

				E_MAGAZINE_OPERATION.PUT:
					CASE uiStep OF
						0:
							IF stRobotStatus.xRotatedToBlank THEN
								Diag.eState := E_MAGAZINE_STATE.NEXT;
							ELSE
								stActiveRobotCommand.eAction := E_ROBOT_ACTION.ROTATE_TO_BLANK;
							END_IF;
						1:
							stActiveRobotCommand.eAction := E_ROBOT_ACTION.MOVE_TO_POINT;
							stActiveRobotCommand.eSetPoint := E_POINT_NAME.MAGAZINE_SAFE;
						2:
							stActiveRobotCommand.eAction := E_ROBOT_ACTION.MOVE_TO_POINT;
							stActiveRobotCommand.eSetPoint := E_POINT_NAME.MAGAZINE_IN_SLOT;
						3: stActiveRobotCommand.eAction := E_ROBOT_ACTION.UNCLAMP_2;
						4:
							stActiveRobotCommand.eAction := E_ROBOT_ACTION.MOVE_TO_POINT;
							stActiveRobotCommand.eSetPoint := E_POINT_NAME.MAGAZINE_SAFE;
					ELSE
						xOperationSequenceComplete := TRUE;
						Diag.eState := E_MAGAZINE_STATE.DONE;
					END_CASE;

				E_MAGAZINE_OPERATION.CHANGE:
					CASE uiStep OF
						0:
							IF (xChangeTakeFirst AND stRobotStatus.xRotatedToDetail)
							OR (NOT xChangeTakeFirst AND stRobotStatus.xRotatedToBlank) THEN
								Diag.eState := E_MAGAZINE_STATE.NEXT;
							ELSIF xChangeTakeFirst THEN
								stActiveRobotCommand.eAction := E_ROBOT_ACTION.ROTATE_TO_DETAIL;
							ELSE
								stActiveRobotCommand.eAction := E_ROBOT_ACTION.ROTATE_TO_BLANK;
							END_IF;
						1:
							stActiveRobotCommand.eAction := E_ROBOT_ACTION.MOVE_TO_POINT;
							stActiveRobotCommand.eSetPoint := E_POINT_NAME.MAGAZINE_SAFE;
						2:
							stActiveRobotCommand.eAction := E_ROBOT_ACTION.MOVE_TO_POINT;
							stActiveRobotCommand.eSetPoint := E_POINT_NAME.MAGAZINE_IN_SLOT;
						3:
							IF xChangeTakeFirst THEN
								stActiveRobotCommand.eAction := E_ROBOT_ACTION.CLAMP_1;
							ELSE
								stActiveRobotCommand.eAction := E_ROBOT_ACTION.UNCLAMP_2;
							END_IF;
						4:
							stActiveRobotCommand.eAction := E_ROBOT_ACTION.MOVE_TO_POINT;
							stActiveRobotCommand.eSetPoint := E_POINT_NAME.MAGAZINE_CHANGE;
						5:
							IF (xChangeTakeFirst AND stRobotStatus.xRotatedToBlank)
							OR (NOT xChangeTakeFirst AND stRobotStatus.xRotatedToDetail) THEN
								Diag.eState := E_MAGAZINE_STATE.NEXT;
							ELSIF xChangeTakeFirst THEN
								stActiveRobotCommand.eAction := E_ROBOT_ACTION.ROTATE_TO_BLANK;
							ELSE
								stActiveRobotCommand.eAction := E_ROBOT_ACTION.ROTATE_TO_DETAIL;
							END_IF;
						6:
							stActiveRobotCommand.eAction := E_ROBOT_ACTION.MOVE_TO_POINT;
							stActiveRobotCommand.eSetPoint := E_POINT_NAME.MAGAZINE_CHANGE;
						7:
							stActiveRobotCommand.eAction := E_ROBOT_ACTION.MOVE_TO_POINT;
							stActiveRobotCommand.eSetPoint := E_POINT_NAME.MAGAZINE_IN_SLOT;
						8:
							IF xChangeTakeFirst THEN
								stActiveRobotCommand.eAction := E_ROBOT_ACTION.UNCLAMP_2;
							ELSE
								stActiveRobotCommand.eAction := E_ROBOT_ACTION.CLAMP_1;
							END_IF;
						9:
							stActiveRobotCommand.eAction := E_ROBOT_ACTION.MOVE_TO_POINT;
							stActiveRobotCommand.eSetPoint := E_POINT_NAME.MAGAZINE_SAFE;
					ELSE
						xOperationSequenceComplete := TRUE;
						Diag.eState := E_MAGAZINE_STATE.DONE;
					END_CASE;

				E_MAGAZINE_OPERATION.RETURN_BLANK:
					CASE uiStep OF
						0:
							IF stRobotStatus.xRotatedToDetail THEN
								Diag.eState := E_MAGAZINE_STATE.NEXT;
							ELSE
								stActiveRobotCommand.eAction := E_ROBOT_ACTION.ROTATE_TO_DETAIL;
							END_IF;
						1:
							stActiveRobotCommand.eAction := E_ROBOT_ACTION.MOVE_TO_POINT;
							stActiveRobotCommand.eSetPoint := E_POINT_NAME.MAGAZINE_SAFE;
						2:
							stActiveRobotCommand.eAction := E_ROBOT_ACTION.MOVE_TO_POINT;
							stActiveRobotCommand.eSetPoint := E_POINT_NAME.MAGAZINE_IN_SLOT;
						3: stActiveRobotCommand.eAction := E_ROBOT_ACTION.UNCLAMP_1;
						4:
							stActiveRobotCommand.eAction := E_ROBOT_ACTION.MOVE_TO_POINT;
							stActiveRobotCommand.eSetPoint := E_POINT_NAME.MAGAZINE_SAFE;
					ELSE
						xOperationSequenceComplete := TRUE;
						Diag.eState := E_MAGAZINE_STATE.DONE;
					END_CASE;
		END_CASE;

		IF Diag.eState = E_MAGAZINE_STATE.PREPARE_STEP THEN
			Diag.eState := E_MAGAZINE_STATE.ROBOT_COMMAND;
		END_IF;

	E_MAGAZINE_STATE.ROBOT_COMMAND:
		Command := stActiveRobotCommand;
		Command.xExecute := TRUE;
		IF stRobotStatus.xBusy THEN
			xRobotCommandStarted := TRUE;
		END_IF;

		IF xStopRequest OR xGlobalError THEN
			Command.xStop := stRobotStatus.xBusy;
			Error.dwErrorActive := Error.dwErrorActive OR ERR_GLOBAL_STOP;
			Diag.eState := E_MAGAZINE_STATE.ERROR;

		ELSIF stRobotStatus.xError THEN
			Error.dwErrorActive := Error.dwErrorActive OR ERR_ROBOT;
			Diag.eState := E_MAGAZINE_STATE.ERROR;

		ELSIF xRobotCommandStarted AND stRobotStatus.xDone THEN
			// Матрица меняется в момент подтверждённого физического переноса,
			// а не после отхода робота и завершения всей составной операции.
			CASE eActualOperation OF
				E_MAGAZINE_OPERATION.TAKE:
					IF (uiStep = UINT#3) AND NOT xTakeSlotCommitted THEN
						xInventoryUpdated := TRUE;
						xInventorySummaryDirty := TRUE;
						stInventory.aSlots[iTakeSlot].xInPosition := FALSE;
						stInventory.aSlots[iTakeSlot].eDetailType := E_DETAIL_TYPE.NONE;
						stInventory.aSlots[iTakeSlot].uiProductType := UINT#0;
						xTakeSlotCommitted := TRUE;
					END_IF;

				E_MAGAZINE_OPERATION.PUT:
					IF (uiStep = UINT#3) AND NOT xPutSlotCommitted THEN
						xInventoryUpdated := TRUE;
						xInventorySummaryDirty := TRUE;
						stInventory.aSlots[iPutSlot].xInPosition := TRUE;
						stInventory.aSlots[iPutSlot].eDetailType := E_DETAIL_TYPE.DETAIL;
						stInventory.aSlots[iPutSlot].uiProductType := uiPutProductType;
						udiProducedPartsTotal := udiProducedPartsTotal + UDINT#1;
						xPutSlotCommitted := TRUE;
					END_IF;

				E_MAGAZINE_OPERATION.CHANGE:
					IF (((uiStep = UINT#3) AND NOT xChangeTakeFirst)
						OR ((uiStep = UINT#8) AND xChangeTakeFirst))
					AND NOT xPutSlotCommitted THEN
						xInventoryUpdated := TRUE;
						xInventorySummaryDirty := TRUE;
						stInventory.aSlots[iPutSlot].xInPosition := TRUE;
						stInventory.aSlots[iPutSlot].eDetailType := E_DETAIL_TYPE.DETAIL;
						stInventory.aSlots[iPutSlot].uiProductType := uiPutProductType;
						udiProducedPartsTotal := udiProducedPartsTotal + UDINT#1;
						xPutSlotCommitted := TRUE;
					ELSIF (((uiStep = UINT#8) AND NOT xChangeTakeFirst)
						OR ((uiStep = UINT#3) AND xChangeTakeFirst))
					AND NOT xTakeSlotCommitted THEN
						xInventoryUpdated := TRUE;
						xInventorySummaryDirty := TRUE;
						stInventory.aSlots[iTakeSlot].xInPosition := FALSE;
						stInventory.aSlots[iTakeSlot].eDetailType := E_DETAIL_TYPE.NONE;
						stInventory.aSlots[iTakeSlot].uiProductType := UINT#0;
						xTakeSlotCommitted := TRUE;
					END_IF;

				E_MAGAZINE_OPERATION.RETURN_BLANK:
					IF (uiStep = UINT#3) AND NOT xPutSlotCommitted THEN
						xFinishedLatched := FALSE;
						xFinishedCondition := FALSE;
						xInventoryUpdated := TRUE;
						xInventorySummaryDirty := TRUE;
						stInventory.aSlots[iPutSlot].xInPosition := TRUE;
						stInventory.aSlots[iPutSlot].eDetailType := E_DETAIL_TYPE.BLANK;
						stInventory.aSlots[iPutSlot].uiProductType := uiPutProductType;
						xPutSlotCommitted := TRUE;
					END_IF;
			END_CASE;
			Diag.eState := E_MAGAZINE_STATE.RELEASE_ROBOT_COMMAND;
		END_IF;

	E_MAGAZINE_STATE.RELEASE_ROBOT_COMMAND:
		IF stRobotStatus.xError THEN
			Error.dwErrorActive := Error.dwErrorActive OR ERR_ROBOT;
			Diag.eState := E_MAGAZINE_STATE.ERROR;
		ELSIF NOT stRobotStatus.xBusy AND NOT stRobotStatus.xDone THEN
			Diag.eState := E_MAGAZINE_STATE.NEXT;
		END_IF;

	E_MAGAZINE_STATE.NEXT:
		uiStep := uiStep + 1;
		Diag.eState := E_MAGAZINE_STATE.PREPARE_STEP;

	E_MAGAZINE_STATE.DONE:
		// Страховочная фиксация нужна только если конечный DONE получен без
		// промежуточного обновления. В штатном ходе слоты уже изменены захватами.
		IF xOperationSequenceComplete
		AND NOT xStopRequest
		AND NOT xGlobalError
		AND NOT xInventoryCommitted THEN
			CASE eActualOperation OF
				E_MAGAZINE_OPERATION.TAKE:
					IF NOT xTakeSlotCommitted THEN
						xInventoryUpdated := TRUE;
						xInventorySummaryDirty := TRUE;
						stInventory.aSlots[iTakeSlot].xInPosition := FALSE;
						stInventory.aSlots[iTakeSlot].eDetailType := E_DETAIL_TYPE.NONE;
						stInventory.aSlots[iTakeSlot].uiProductType := UINT#0;
						xTakeSlotCommitted := TRUE;
					END_IF;
				E_MAGAZINE_OPERATION.PUT:
					IF NOT xPutSlotCommitted THEN
						xInventoryUpdated := TRUE;
						xInventorySummaryDirty := TRUE;
						stInventory.aSlots[iPutSlot].xInPosition := TRUE;
						stInventory.aSlots[iPutSlot].eDetailType := E_DETAIL_TYPE.DETAIL;
						stInventory.aSlots[iPutSlot].uiProductType := uiPutProductType;
						udiProducedPartsTotal := udiProducedPartsTotal + UDINT#1;
						xPutSlotCommitted := TRUE;
					END_IF;
				E_MAGAZINE_OPERATION.CHANGE:
					// Для обмена в одном слоте сначала отражаем изъятие. Уже
					// подтверждённую укладку нельзя затереть страховочной фиксацией.
					IF NOT xTakeSlotCommitted THEN
						IF NOT xChangeTakeFirst OR NOT xPutSlotCommitted THEN
							xInventoryUpdated := TRUE;
							xInventorySummaryDirty := TRUE;
							stInventory.aSlots[iTakeSlot].xInPosition := FALSE;
							stInventory.aSlots[iTakeSlot].eDetailType := E_DETAIL_TYPE.NONE;
							stInventory.aSlots[iTakeSlot].uiProductType := UINT#0;
						END_IF;
						xTakeSlotCommitted := TRUE;
					END_IF;
					IF NOT xPutSlotCommitted THEN
						xInventoryUpdated := TRUE;
						xInventorySummaryDirty := TRUE;
						stInventory.aSlots[iPutSlot].xInPosition := TRUE;
						stInventory.aSlots[iPutSlot].eDetailType := E_DETAIL_TYPE.DETAIL;
						stInventory.aSlots[iPutSlot].uiProductType := uiPutProductType;
						udiProducedPartsTotal := udiProducedPartsTotal + UDINT#1;
						xPutSlotCommitted := TRUE;
					END_IF;
				E_MAGAZINE_OPERATION.RETURN_BLANK:
					IF NOT xPutSlotCommitted THEN
						xFinishedLatched := FALSE;
						xFinishedCondition := FALSE;
						xInventoryUpdated := TRUE;
						xInventorySummaryDirty := TRUE;
						stInventory.aSlots[iPutSlot].xInPosition := TRUE;
						stInventory.aSlots[iPutSlot].eDetailType := E_DETAIL_TYPE.BLANK;
						stInventory.aSlots[iPutSlot].uiProductType := uiPutProductType;
						xPutSlotCommitted := TRUE;
					END_IF;
			END_CASE;
			xInventoryCommitted := TRUE;
		END_IF;
		IF NOT xExecuteRequest THEN
			eActualOperation := E_MAGAZINE_OPERATION.NONE;
			IF xDisableRequest
			AND NOT xRobotInMagazineContext THEN
				Diag.eState := E_MAGAZINE_STATE.DISABLED;
			ELSE
				Diag.eState := E_MAGAZINE_STATE.IDLE;
			END_IF;
		END_IF;

	E_MAGAZINE_STATE.ERROR:
		IF (rtReset.Q OR xRobotResetAttemptReady)
		AND NOT xResetCancel
		AND NOT xIoManual
		AND NOT xExecuteRequest
		AND NOT xStopRequest
		AND NOT FaultStatus.xBusy
		AND NOT xGlobalError
		AND xRobotResetDependencyReady THEN
			IF xRobotResetDependencyRequired AND stRobotStatus.xError AND NOT xRobotResetAttemptReady THEN
				// Не очищаем каскад заранее: робот ещё восстанавливает Motion.
				// Без его принятой попытки местный Reset ничего не повторяет.
				xRobotResetCoordinated := TRUE;
				udiRobotResetAttempt := RobotResetRecovery.udiAttempt + UDINT#1;
				IF udiRobotResetAttempt = UDINT#0 THEN udiRobotResetAttempt := UDINT#1; END_IF;
			ELSE
				Error.dwErrorLast := Error.dwErrorActive;
				Error.dwErrorActive := DWORD#0;
				eActualOperation := E_MAGAZINE_OPERATION.NONE;
				Diag.eState := E_MAGAZINE_STATE.DISABLED;
			END_IF;
		END_IF;
END_CASE;

// Класс реакции не размазывается по CASE. Первичная причина остаётся в своей
// маске, а контекст конкретного магазина хранится до принятого сброса.
IF (Diag.eState = E_MAGAZINE_STATE.ERROR)
AND NOT xFaultContextCaptured THEN
	xRobotInMagazineAtFault := xRobotInMagazineContext;
	xFaultContextCaptured := TRUE;
ELSIF Diag.eState <> E_MAGAZINE_STATE.ERROR THEN
	xRobotInMagazineAtFault := FALSE;
	xFaultContextCaptured := FALSE;
END_IF;

xRobotStopRequired := NOT xGlobalError
	AND (
		((Error.dwErrorActive AND ERR_ROBOT) <> DWORD#0)
		OR (((Error.dwErrorActive AND MASK_EQUIPMENT_ERROR) <> DWORD#0)
			AND xRobotInMagazineAtFault)
	);

// Физический Stop нужен только занятому роботу. При неподвижном роботе внутри
// магазина FB_ROBOT получит зависимую ошибку без пустой команды остановки.
IF (Diag.eState = E_MAGAZINE_STATE.ERROR)
AND xRobotStopRequired
AND stRobotStatus.xBusy THEN
	Command := stActiveRobotCommand;
	Command.xExecute := TRUE;
	Command.xStop := TRUE;
END_IF;

// ERROR технологически отключает магазин немедленно, но причина остаётся
// защёлкнутой до разрешённого Reset.
Status.xEnabled := (Diag.eState <> E_MAGAZINE_STATE.DISABLED)
	AND (Diag.eState <> E_MAGAZINE_STATE.ERROR);
Status.xDisablePending := xDisableRequest AND Status.xEnabled;
Status.xPowerAllowed := Status.xEnabled OR Status.xEnableSequenceAllowed;
Status.xFillAllowed := (iActiveSlotCount > SINT#0) AND Status.xEditAllowed;
Status.xClearAllowed := Status.xEditAllowed;
Status.xReady := xMechanismReady AND  (Diag.eState = E_MAGAZINE_STATE.IDLE)
	AND xRobotCanWorkWithMagazine
	AND (Error.dwErrorActive = DWORD#0);
Status.xBusy := (Diag.eState <> E_MAGAZINE_STATE.DISABLED)
	AND (Diag.eState <> E_MAGAZINE_STATE.IDLE)
	AND (Diag.eState <> E_MAGAZINE_STATE.DONE)
	AND (Diag.eState <> E_MAGAZINE_STATE.ERROR);
Status.xDone := Diag.eState = E_MAGAZINE_STATE.DONE;
Status.xError := Diag.eState = E_MAGAZINE_STATE.ERROR;
Status.xRobotStopRequired := xRobotStopRequired;
Status.udiProducedPartsTotal := udiProducedPartsTotal;
Status.uiMagazineId := uiMagazineId;
Status.eGrantedOperation := eGrantedOperation;
Status.eActualOperation := eActualOperation;
Status.iSelectedBlank := iTakeSlot;
Status.iSelectedFreeSlot := iPutSlot;
// Разовая доработка палеты завершена: чужой груз/станок не возвращает её
// в планирование. Защёлку снимает только смена банка или правка его содержимого.
xFinishedLatched := xFinishedLatched OR (xFinishedCondition AND NOT Status.xBusy);
Status.xFinished := xFinishedLatched;
Error.dwAlarmActive := Error.dwErrorActive;

IF Error.dwErrorActive <> DWORD#0 THEN
	Error.dwErrorLast := Error.dwErrorActive;
END_IF;

Error.stErrorActive := UpdateErrorView(dwError := Error.dwErrorActive);
Error.stErrorLast := UpdateErrorView(dwError := Error.dwErrorLast);
FaultStatus.xResetAllowed := Status.xError
	AND NOT xRobotResetCoordinated
	AND NOT xResetCancel
	AND NOT xIoManual
	AND NOT FaultStatus.xBusy
	AND NOT xExecuteRequest
	AND NOT xStopRequest
	AND NOT xGlobalError
	AND xRobotResetDependencyReady;

// Подтверждение захвата/укладки обновляет сводку в том же скане.
// В ожидании повторный проход не нужен; выбор операции сохраняет прежний порядок.
IF xInventorySummaryDirty THEN
    UpdateTypeStatus(stMagazineInventory := stInventory);
END_IF;

(* ---- FB_MOTION_MANAGER.st ---- *)
FUNCTION_BLOCK FB_MOTION_MANAGER
VAR_INPUT
	stPoint : ARRAY [0..GVL_POINT.iPointNumber] OF ST_POINT; // Глобальная таблица точек
	xReset  : BOOL; // Сброс ошибок менеджера движения
	FaultRequest : ST_POINT_FAULT_REQUEST; // Диагностические ошибки проверки точки
	xSpeedFactorOverride : BOOL; // Для отдельной проверки точки с телефона
	lrSpeedFactorOverride : LREAL; // 0.001..1.0, применяется вместо SpeedFactor точки
	lrAccelerationFactor : LREAL := 1.0; // Единый предел разгона/торможения группы 0.01..1.0
	lrJerkFactor : LREAL := 1.0; // Плавность групповой траектории 0.01..1.0
END_VAR
VAR_OUTPUT
	FaultStatus : ST_FAULT_INJECTION_STATUS; // Состояние инжектора проверки точки
END_VAR
VAR
	curPoint      : ST_POINT; // Координаты выбранной точки
	curPointName  : E_POINT_NAME; // Имя выбранной точки
	fbPointManager: FB_POINT_MANAGER; // Проверка координат и скорости точки
	fbPointFaultInjector : FB_POINT_FAULT_INJECTOR; // Безопасная подмена проверяемой точки
	rtReset       : R_TRIG; // Фронт команды сброса менеджера движения
	xFaultAllowed : BOOL; // Менеджер готов к синтетической проверке без движения
	xGroupMotionStarted : BOOL; // Группа приняла движение, ожидание запуска завершено
	tonMotionStart : TON; // Общий предел проверки точки и старта группы
END_VAR
VAR CONSTANT
	ERR_POINT_INVALID : DWORD := DWORD#16#0000_0001; // Недопустимая точка
	ERR_GROUP         : DWORD := DWORD#16#0000_0002; // Ошибка группы осей
	ERR_GLOBAL_STOP   : DWORD := DWORD#16#0000_0004; // Глобальная ошибка ячейки
	ERR_START_TIMEOUT : DWORD := DWORD#16#0000_0008; // Проверка/запуск группы не завершены вовремя
	WRN_RESET_GLOBAL_ERROR : UINT := 1; // Глобальная ошибка ещё активна
	WRN_SIM_ERROR_NOT_ALLOWED : UINT := 2; // Тестовая проверка запрещена текущим состоянием
END_VAR
VAR_IN_OUT
	stMotionManager : ST_MOTION_MANAGER; // Команды, статусы и диагностика менеджера движения
	GroupData       : ST_AXIS_GROUP; // Команды, статусы и диагностика группы XYZ
	stPointManager  : ST_POINT_MANAGER; // Команды, статусы и диагностика проверки точки
END_VAR

// --- BEGIN IMPLEMENTATION ---

xFaultAllowed := (stMotionManager.Diag.eState = E_MOTION_MANAGER_STATE.IDLE)
	AND NOT stMotionManager.Command.xExecute
	AND NOT stMotionManager.Command.xGlobalError
	AND (stMotionManager.Error.dwErrorActive = DWORD#0)
	AND NOT GroupData.Status.xLocalError
	AND NOT GroupData.Command.xMoveDirect
	AND NOT GroupData.Command.xMoveLinear;

fbPointFaultInjector(
	Request := FaultRequest,
	xOwnerAllowed := xFaultAllowed,
	xComplete := stMotionManager.Diag.eState = E_MOTION_MANAGER_STATE.ERROR,
	PointRaw := stPoint[E_POINT_NAME.MAGAZINE_DETAIL]
);
FaultStatus := fbPointFaultInjector.Status;

IF fbPointFaultInjector.Status.xRejected THEN
	stPointManager.Diag.stWarning.uiCode := WRN_SIM_ERROR_NOT_ALLOWED;
	stPointManager.Diag.stWarning.udiSequence := stPointManager.Diag.stWarning.udiSequence + UDINT#1;
	IF stPointManager.Diag.stWarning.udiSequence = UDINT#0 THEN
		stPointManager.Diag.stWarning.udiSequence := UDINT#1;
	END_IF;
END_IF;

IF fbPointFaultInjector.xExecute THEN
	curPoint := fbPointFaultInjector.Point;
	curPointName := E_POINT_NAME.NONE;
END_IF;

// Рабочая точка должна быть защёлкнута до вызова FB_POINT_MANAGER. Иначе при
// переходе в VALIDATE менеджер точек видит curPoint от предыдущей команды
// (или нулевой ST_POINT при первом проходе), потому что прежняя запись
// выполнялась ниже вызова FB_POINT_MANAGER в CASE VALIDATE.
IF (stMotionManager.Diag.eState = E_MOTION_MANAGER_STATE.VALIDATE)
AND NOT fbPointFaultInjector.xExecute THEN

	curPoint := stPoint[stMotionManager.Command.eTargetPoint];
	curPointName := stMotionManager.Command.eTargetPoint;
END_IF;

fbPointManager(
			stPointManager := stPointManager,
			stPoint := curPoint
		);

stMotionManager.Status.xBusy := FALSE;
stMotionManager.Status.xDone := FALSE;
stMotionManager.Status.xError := FALSE;
stMotionManager.Status.xReady:= FALSE;
stMotionManager.Command.xReset := xReset;
rtReset(CLK := xReset);

IF rtReset.Q
AND (stMotionManager.Diag.eState = E_MOTION_MANAGER_STATE.ERROR)
AND stMotionManager.Command.xGlobalError THEN
	stMotionManager.Diag.stWarning.uiCode := WRN_RESET_GLOBAL_ERROR;
	stMotionManager.Diag.stWarning.udiSequence := stMotionManager.Diag.stWarning.udiSequence + UDINT#1;
	IF stMotionManager.Diag.stWarning.udiSequence = UDINT#0 THEN
		stMotionManager.Diag.stWarning.udiSequence := UDINT#1;
	END_IF;
END_IF;

IF (stMotionManager.Diag.eState = E_MOTION_MANAGER_STATE.MOTION_SIM)
AND ((GroupData.Diag.iStep = E_AXIS_GROUP_STATE.MOVING_DIRECT)
	OR (GroupData.Status.xMoveDirectDone AND GroupData.Command.xMoveDirect)) THEN
	xGroupMotionStarted := TRUE;
END_IF;
tonMotionStart(
	IN := (stMotionManager.Diag.eState = E_MOTION_MANAGER_STATE.VALIDATE)
		OR ((stMotionManager.Diag.eState = E_MOTION_MANAGER_STATE.MOTION_SIM)
			AND NOT xGroupMotionStarted),
	PT := GroupData.Timeouts.tGroupTimeout
);

// Stop должен отменять ещё не запущенную команду и завершённую команду,
// ожидающую освобождения. Проверка точки тоже получает спад Execute.
IF stMotionManager.Command.xGlobalError THEN
	stPointManager.Command.xExecute := FALSE;
	GroupData.Command.xMoveDirect := FALSE;
	GroupData.Command.xMoveLinear := FALSE;
	stMotionManager.Error.dwErrorActive := stMotionManager.Error.dwErrorActive OR ERR_GLOBAL_STOP;
	stMotionManager.Diag.eState := E_MOTION_MANAGER_STATE.ERROR;
ELSIF stMotionManager.Command.xStop
AND (stMotionManager.Diag.eState <> E_MOTION_MANAGER_STATE.ERROR) THEN
	stPointManager.Command.xExecute := FALSE;
	GroupData.Command.xMoveDirect := FALSE;
	GroupData.Command.xMoveLinear := FALSE;
	xGroupMotionStarted := FALSE;
	stMotionManager.Diag.eState := E_MOTION_MANAGER_STATE.IDLE;
ELSIF tonMotionStart.Q THEN
	stPointManager.Command.xExecute := FALSE;
	GroupData.Command.xMoveDirect := FALSE;
	GroupData.Command.xMoveLinear := FALSE;
	stMotionManager.Error.dwErrorActive := stMotionManager.Error.dwErrorActive OR ERR_START_TIMEOUT;
	stMotionManager.Diag.eState := E_MOTION_MANAGER_STATE.ERROR;
END_IF;

CASE stMotionManager.Diag.eState OF
	// --------------------------------------------------
	E_MOTION_MANAGER_STATE.IDLE:
	// --------------------------------------------------
		// Менеджер является единственным владельцем команд движения группы.
		// После завершения или сброса не оставляем уровень Execute защёлкнутым.
		GroupData.Command.xMoveDirect := FALSE;
		GroupData.Command.xMoveLinear := FALSE;
		xGroupMotionStarted := FALSE;
		stMotionManager.Status.xReady:= TRUE;
		IF (stMotionManager.Command.xExecute OR fbPointFaultInjector.xExecute)
		AND NOT stMotionManager.Command.xGlobalError
		AND NOT stMotionManager.Command.xStop THEN
			stMotionManager.Status.xBusy := TRUE;
			stMotionManager.Diag.eState := E_MOTION_MANAGER_STATE.VALIDATE;
		ELSIF stMotionManager.Command.xGlobalError THEN
			stMotionManager.Error.dwErrorActive := stMotionManager.Error.dwErrorActive OR ERR_GLOBAL_STOP;
			stMotionManager.Diag.eState := E_MOTION_MANAGER_STATE.ERROR;
		END_IF;

	// --------------------------------------------------
	E_MOTION_MANAGER_STATE.VALIDATE:
	// --------------------------------------------------
		stMotionManager.Status.xBusy := TRUE;
		stPointManager.Command.xExecute := TRUE;

		IF stPointManager.Status.xDone AND NOT stPointManager.Status.xInvalid THEN
			stPointManager.Command.xExecute := FALSE;
			IF stMotionManager.Command.xMode THEN
				stMotionManager.Diag.eState := 	E_MOTION_MANAGER_STATE.MOTION_MODBUS;
			ELSE
				stMotionManager.Diag.eState := 	E_MOTION_MANAGER_STATE.MOTION_SIM;
			END_IF;
		ELSIF stPointManager.Status.xDone AND stPointManager.Status.xInvalid THEN
			stPointManager.Command.xExecute := FALSE;
			stMotionManager.Error.dwErrorActive := stMotionManager.Error.dwErrorActive OR ERR_POINT_INVALID;
			stMotionManager.Diag.eState := 	E_MOTION_MANAGER_STATE.ERROR;
		END_IF;

	// --------------------------------------------------
	E_MOTION_MANAGER_STATE.MOTION_SIM:
	// --------------------------------------------------

		stMotionManager.Status.xBusy := TRUE;

		GroupData.MotionParam.lrX := curPoint.X;
		GroupData.MotionParam.lrY := curPoint.Y;
		GroupData.MotionParam.lrZ := curPoint.Z;
		IF xSpeedFactorOverride THEN
			GroupData.MotionParam.VelFactor := LIMIT(0.001, lrSpeedFactorOverride, 1.0);
		ELSE
			GroupData.MotionParam.VelFactor := curPoint.SpeedFactor;
		END_IF;
		// У группы SoftMotion один AccFactor для обеих сторон профиля. PLC передаёт
		// сюда более строгий из глобальных процентов разгона и торможения.
		GroupData.MotionParam.AccFactor := LIMIT(0.01, lrAccelerationFactor, 1.0);
		GroupData.MotionParam.JerkFactor := LIMIT(0.01, lrJerkFactor, 1.0);
		IF GroupData.Diag.iStep = E_AXIS_GROUP_STATE.READY
		AND NOT GroupData.Command.xMoveDirect
		AND NOT stMotionManager.Command.xGlobalError
		AND NOT stMotionManager.Command.xStop THEN
			GroupData.Command.xMoveDirect := TRUE;
		END_IF;

		IF stMotionManager.Command.xStop THEN
			GroupData.Command.xMoveDirect := FALSE;
			GroupData.Command.xMoveLinear := FALSE;
			stMotionManager.Status.xBusy := FALSE;
			stMotionManager.Diag.eState := E_MOTION_MANAGER_STATE.IDLE;
		ELSIF GroupData.Status.xMoveDirectDone AND GroupData.Command.xMoveDirect THEN
			GroupData.Command.xMoveDirect := FALSE;
			stMotionManager.Status.eCurrentPoint := curPointName;
			stMotionManager.Diag.eState := 	E_MOTION_MANAGER_STATE.DONE;
		ELSIF GroupData.Diag.iStep = E_AXIS_GROUP_STATE.ERROR OR stMotionManager.Command.xGlobalError  THEN
			GroupData.Command.xMoveDirect := FALSE;
			GroupData.Command.xMoveLinear := FALSE;
			IF GroupData.Diag.iStep = E_AXIS_GROUP_STATE.ERROR THEN
				stMotionManager.Error.dwErrorActive := stMotionManager.Error.dwErrorActive OR ERR_GROUP;
			END_IF;
			IF stMotionManager.Command.xGlobalError THEN
				stMotionManager.Error.dwErrorActive := stMotionManager.Error.dwErrorActive OR ERR_GLOBAL_STOP;
			END_IF;
			stMotionManager.Diag.eState := 	E_MOTION_MANAGER_STATE.ERROR;
		END_IF;

	// --------------------------------------------------
	E_MOTION_MANAGER_STATE.ERROR:
	// --------------------------------------------------
		GroupData.Command.xMoveDirect := FALSE;
		GroupData.Command.xMoveLinear := FALSE;
		stMotionManager.Status.xError := TRUE;
		IF NOT stMotionManager.Command.xGlobalError AND stMotionManager.Command.xReset THEN
			stMotionManager.Error.dwErrorLast := stMotionManager.Error.dwErrorActive;
			stMotionManager.Error.dwErrorActive := DWORD#0;
			stMotionManager.Status.xError := FALSE;
			stMotionManager.Diag.eState := 	E_MOTION_MANAGER_STATE.IDLE;
		END_IF;

	// --------------------------------------------------
	E_MOTION_MANAGER_STATE.DONE:
	// --------------------------------------------------
		stMotionManager.Status.xBusy := FALSE;
		stMotionManager.Status.xDone := TRUE;
		IF NOT stMotionManager.Command.xExecute THEN
			stMotionManager.Diag.eState := 	E_MOTION_MANAGER_STATE.IDLE;
		END_IF;
	END_CASE;

// Журнал отражает состояние каждого FB, включая каскадные ошибки зависимостей.
stMotionManager.Error.dwAlarmActive := stMotionManager.Error.dwErrorActive;

stMotionManager.Error.stErrorActive := UpdateErrorView(
	dwError := stMotionManager.Error.dwErrorActive
);
stMotionManager.Error.stErrorLast := UpdateErrorView(
	dwError := stMotionManager.Error.dwErrorLast
);
FaultStatus.xResetAllowed := stMotionManager.Status.xError
	AND NOT FaultStatus.xBusy;

(* ---- FB_POINT_MANAGER.st ---- *)
FUNCTION_BLOCK FB_POINT_MANAGER
VAR_INPUT
	stPoint : ST_POINT; // Проверяемая точка
END_VAR
VAR_OUTPUT
END_VAR
VAR
END_VAR
VAR_IN_OUT
	stPointManager : ST_POINT_MANAGER; // Команды, статусы и диагностика проверки точки
END_VAR
VAR CONSTANT
	X_OUT_OF_LIMIT : DWORD := 1; // Координата X вне допустимых границ
	Y_OUT_OF_LIMIT : DWORD := 2; // Координата Y вне допустимых границ
	Z_OUT_OF_LIMIT : DWORD := 4; // Координата Z вне допустимых границ
	INVALID_VEL    : DWORD := 8; // Недопустимый коэффициент скорости
	X_LIMIT_CONFIG_INVALID : DWORD := 16; // Software limits оси X недоступны или некорректны
	Y_LIMIT_CONFIG_INVALID : DWORD := 32; // Software limits оси Y недоступны или некорректны
	Z_LIMIT_CONFIG_INVALID : DWORD := 64; // Software limits оси Z недоступны или некорректны
	POINT_NOT_CONFIGURED : DWORD := 128; // Инженерная точка не подтверждена редактором
END_VAR

// --- BEGIN IMPLEMENTATION ---

stPointManager.Status.xBusy := FALSE;
stPointManager.Status.xDone := FALSE;
stPointManager.Status.xInvalid := FALSE;

CASE stPointManager.Diag.eState OF
	// --------------------------------------------------
	E_POINT_MANAGER_STATE.IDLE:
	// --------------------------------------------------
		stPointManager.Error.dwErrorActive := DWORD#0;
		IF stPointManager.Command.xExecute THEN
			stPointManager.Status.xBusy := TRUE;
			stPointManager.Diag.eState := E_POINT_MANAGER_STATE.CHECK_ZONE;
		END_IF

	// --------------------------------------------------
	E_POINT_MANAGER_STATE.CHECK_ZONE:
	// --------------------------------------------------
		stPointManager.Status.xBusy := TRUE;
		IF NOT stPoint.xConfigured THEN
			stPointManager.Error.dwErrorActive :=
				stPointManager.Error.dwErrorActive OR POINT_NOT_CONFIGURED;
		END_IF

		IF NOT stPointManager.Diag.xXLimitValid
		OR NOT stPointManager.Diag.xYLimitValid
		OR NOT stPointManager.Diag.xZLimitValid THEN
			// Без достоверных активных SoftMotion limits движение к точке запрещается.
			// Статический резервный диапазон здесь намеренно не применяется.
			IF NOT stPointManager.Diag.xXLimitValid THEN
				stPointManager.Error.dwErrorActive :=
					stPointManager.Error.dwErrorActive OR X_LIMIT_CONFIG_INVALID;
			END_IF
			IF NOT stPointManager.Diag.xYLimitValid THEN
				stPointManager.Error.dwErrorActive :=
					stPointManager.Error.dwErrorActive OR Y_LIMIT_CONFIG_INVALID;
			END_IF
			IF NOT stPointManager.Diag.xZLimitValid THEN
				stPointManager.Error.dwErrorActive :=
					stPointManager.Error.dwErrorActive OR Z_LIMIT_CONFIG_INVALID;
			END_IF
		ELSE
			IF NOT ((stPointManager.Diag.lrX_MinLimit <= stPoint.X) AND (stPoint.X <= stPointManager.Diag.lrX_MaxLimit)) THEN
				stPointManager.Error.dwErrorActive := stPointManager.Error.dwErrorActive OR X_OUT_OF_LIMIT;
			END_IF

			IF NOT ((stPointManager.Diag.lrY_MinLimit <= stPoint.Y) AND (stPoint.Y <= stPointManager.Diag.lrY_MaxLimit)) THEN
				stPointManager.Error.dwErrorActive := stPointManager.Error.dwErrorActive OR Y_OUT_OF_LIMIT;
			END_IF

			IF NOT ((stPointManager.Diag.lrZ_MinLimit <= stPoint.Z) AND (stPoint.Z <= stPointManager.Diag.lrZ_MaxLimit)) THEN
				stPointManager.Error.dwErrorActive := stPointManager.Error.dwErrorActive OR Z_OUT_OF_LIMIT;
			END_IF
		END_IF

		stPointManager.Diag.eState := E_POINT_MANAGER_STATE.CHECK_VEL_FACTOR;

	// --------------------------------------------------
	E_POINT_MANAGER_STATE.CHECK_VEL_FACTOR:
	// --------------------------------------------------
		stPointManager.Status.xBusy := TRUE;

		IF  NOT ((0.1 < stPoint.SpeedFactor) AND(stPoint.SpeedFactor <= 1.0))  THEN
			stPointManager.Error.dwErrorActive := stPointManager.Error.dwErrorActive OR INVALID_VEL;
		END_IF

		stPointManager.Diag.eState := E_POINT_MANAGER_STATE.CHECK_ALL;

	// --------------------------------------------------
	E_POINT_MANAGER_STATE.CHECK_ALL:
	// --------------------------------------------------
		stPointManager.Status.xDone := TRUE;
		stPointManager.Status.xBusy := FALSE;
		IF stPointManager.Error.dwErrorActive <> DWORD#0 THEN
			stPointManager.Status.xInvalid := TRUE;
			stPointManager.Error.dwErrorLast := stPointManager.Error.dwErrorActive;
		ELSE
			stPointManager.Status.xInvalid := FALSE;
		END_IF

		IF NOT stPointManager.Command.xExecute THEN
			stPointManager.Diag.eState := E_POINT_MANAGER_STATE.IDLE;
		END_IF

END_CASE

stPointManager.Error.dwAlarmActive := stPointManager.Error.dwErrorActive;

stPointManager.Error.stErrorActive := UpdateErrorView(
	dwError := stPointManager.Error.dwErrorActive
);
stPointManager.Error.stErrorLast := UpdateErrorView(
	dwError := stPointManager.Error.dwErrorLast
);
